  local PSE_WA_1 = p[ 0.000,-0.400, 0.300, 0.000, 0.000, 0.000]
  local PSE_WA_2 = p[-0.300,-0.300, 0.300, 0.000, 0.000, d2r(-90)]
  local PSE_WA_3 = p[-0.300, 0.300, 0.300, 0.000, 0.000, d2r(-135)]
  local PSE_WA_4 = p[ 0.300, 0.300, 0.300, 0.000, 0.000, d2r(135)]
  local PSE_WA_5 = p[ 0.300,-0.300, 0.300, 0.000, 0.000, d2r(90)]
  local PSE_WA_6 = p[ 0.000,-0.600, 0.300, 0.000, 0.000, 0.000]       # reserved
  local PSE_WA_7 = p[ 0.000, 0.000, 0.000, 0.000, 0.000, 0.000]       # reserved
  local PSE_WA_8 = p[ 0.000, 0.000, 0.000, 0.000, 0.000, 0.000]       # reserved
  local PSE_WA_9 = p[ 0.000, 0.000, 0.000, 0.000, 0.000, 0.000]       # reserved
  local PSE_WA_10 = p[ 0.000, 0.000, 0.000, 0.000, 0.000, 0.000]      # reserved

  local JNT_HOME = [-1.22921,-1.29807,-1.79972,-1.6152, 1.57367, 3.48142]
  local JNT_STANDARD_C1 = [ 1.57,-1.57, 1.57,-1.57,-1.57,0]
  local JNT_STANDARD_C2 = [-1.57,-1.57,-1.57,-1.57, 1.57,0]
  local YAW_MIN_DEG = -110
  local YAW_MAX_DEG = 110
  local DISTANCE_TO_CLEARANCE = 0.300
  local RADIUS_HELPER_POSES = 0.300
  local RADIUS_TRANSITION_POSES = 0.400
  local workareas = [WORKAREA_1, WORKAREA_2, WORKAREA_3, WORKAREA_4, WORKAREA_5, WORKAREA_6, WORKAREA_7, WORKAREA_8, WORKAREA_9, WORKAREA_10]
  local poses = [PSE_WA_1, PSE_WA_2, PSE_WA_3, PSE_WA_4, PSE_WA_5, PSE_WA_6, PSE_WA_7, PSE_WA_8, PSE_WA_9, PSE_WA_10]

  ######################### end of adjustment #########################

  local pi = 3.14159265
  local axis_config_current = 0
  local axis_config_new = 0
  local workarea_current = 0
  local workarea_new = 0
  global reverse_rotation = False
  local pose_start = struct(crt = p[0,0,0,0,0,0], jnt = [0,0,0,0,0,0], q = [0,0,0,0,0,0], yaw_too_base = 0.0)
  local pose_help = struct(crt = p[0,0,0,0,0,0], jnt = [0,0,0,0,0,0], q = [0,0,0,0,0,0], yaw_too_base = 0.0)
  local pose_target = struct(crt = p[0,0,0,0,0,0], jnt = [0,0,0,0,0,0], q = [0,0,0,0,0,0], yaw_too_base = 0.0)
  local pose = struct(crt = p[0,0,0,0,0,0], jnt = [0,0,0,0,0,0], q = [0,0,0,0,0,0], yaw_too_base = 0.0)

  def get_tool_free_pose(pose_ref=get_actual_tcp_pose(), dir=[0,0,0], move_in_base_frame=False):
      # get a recovery pose
      # dir is providing the direction and distance in X, Y and Z
      # if 'move_in_base_frame' is set, dir will be interpreted as absolute values for a movement in base frame

      local pose_target = pose_ref
      local i = 0

      if (move_in_base_frame):
          while (i<3):
              # move only,
              # if the demanded position is bigger than zero and the current position is below the demanded one or
              # if the demanded position is smaller than zero and the current position is above the demanded one
              if ((dir[i]>0 and pose_ref[i]<dir[i]) or (dir[i]<0 and pose_ref[i]>dir[i])):
                  pose_target[i] = dir[i]
              end
              i = i + 1
          end
      else:
          pose_target = pose_trans(pose_ref, p[dir[0], dir[1], dir[2], 0, 0, 0])
      end

      return pose_target
  end

  def check_workarea(reference_pose):
      # the actual TCP position is compared to predefined areas (cubic) to determine in which area the robot arm is
      # a workarea is defined as a list of coordinates, where the first 3 values are X, Y, and Z with the smallest values and
      # the next 3 values specify X, Y and Z for the biggest values

      local data_size = size(workareas)
      local i = 0
      local size_workarea = p[0,0,0,0,0,0]
      local pose_workarea = p[0,0,0,0,0,0]

      while (i < data_size[0]):
          pose_workarea = pose_trans(inv(p[workareas[i, 0], workareas[i, 1], workareas[i, 2], 0, 0, 0]), reference_pose)
          size_workarea = pose_sub(p[workareas[i, 3], workareas[i, 4], workareas[i, 5], 0, 0, 0], p[workareas[i, 0], workareas[i, 1], workareas[i, 2], 0, 0, 0])
          if  ((pose_workarea[0]>0 and pose_workarea[0]<size_workarea[0]) and
              (pose_workarea[1]>0 and pose_workarea[1]<size_workarea[1]) and
              (pose_workarea[2]>0 and pose_workarea[2]<size_workarea[2])):
              return i + 1
          end
          i = i + 1
      end
      return 0
  end

  def check_current_axis_config():
      # function determnines, if the arm is oriented in one or the other configuration.
      # it means, that the ellbow joint is flipped and so are the wrist joints.

      local jnt_current = get_actual_joint_positions()

      # ellbow has positiv angle
      if (jnt_current[2]> 0):
          return 1
      # ellbow has negativ angle
      elif (jnt_current[2]< 0):
          return 2
      # angle is 0
      else:
          return 0
      end
  end

  def switch_axis_config(axis_config):
      # function to switch betwwen the axis configuration 1 and 2.

      if (axis_config == 1):
          return 2
      elif (axis_config ==2):
          return 1
      end
  end

  def get_transition_pose_by_workarea(workarea, axis_config):
      # get the correspondig pose from the list of poses

      pose.crt = poses[workarea-1]
      pose.yaw_too_base = get_yaw_too_base(pose.crt)
      pose.q = get_actual_joint_positions()

      if get_inverse_kin_has_solution(pose.crt, qnear=pose.q):
          pose.jnt = get_inverse_kin(pose.crt, qnear=pose.q)
      else:
          popup("no solution found for the transition pose", blocking= True)
      end

      return pose
  end

  def get_transition_pose_by_reference_pose(ref, radius, axis_config):
      # get the correspondig pose from the list of poses

      pose.yaw_too_base = get_yaw_too_base(ref)
      pose.q = get_actual_joint_positions()

      # get coordinates of the circle with the same angle as the given pose to the
      if ref == p[0,0,0,0,0,0]:
          pose.q = JNT_HOME
          pose.jnt = JNT_HOME
          pose.crt = get_forward_kin(pose.jnt)
          return pose
      else:
          pose.crt = p[
              radius * cos(pose.yaw_too_base-pi/2),
              radius * sin(pose.yaw_too_base-pi/2),
              DISTANCE_TO_CLEARANCE,
              0,
              0,
              pose.yaw_too_base + get_locked_yaw()]
      end

      if get_inverse_kin_has_solution(pose.crt, qnear=pose.q):
          pose.jnt = get_inverse_kin(pose.crt, qnear=pose.q)
      else:
          popup("no solution found for the transition pose", blocking= True)
      end

      return pose
  end

  def get_transition_pose_by_yaw(yaw, radius, axis_config):

      pose.yaw_too_base = yaw
      pose.q = get_actual_joint_positions()
      pose.crt = p[
          radius * cos(yaw-pi/2),
          radius * sin(yaw-pi/2),
          DISTANCE_TO_CLEARANCE,
          0,
          0,
          yaw + get_locked_yaw()]

      if get_inverse_kin_has_solution(pose.crt, qnear=pose.q):
          pose.jnt = get_inverse_kin(pose.crt, qnear=pose.q)
      else:
          popup("no solution found for the transition pose", blocking= True)
      end

      return pose
  end

  def get_rounded_mm(value):
      if (value < 0):
          return ceil(value*1000)
      elif (value >= 0):
          return floor(value*1000)
      end
  end

  def get_yaw_too_base(pose):
      # get the yaw relative to the base frame
      local pose_x_mm = 0
      local pose_y_mm = 0
      local yaw = 0

      pose_x_mm = get_rounded_mm(pose[0])
      pose_y_mm = get_rounded_mm(pose[1])

      if (pose_x_mm == 0 and pose_y_mm < 0):
          yaw = 0
      elif (pose_x_mm == 0 and pose_y_mm > 0):
          yaw = pi
      elif (pose_x_mm < 0 and pose_y_mm == 0):
          yaw = -pi/2
      elif (pose_x_mm > 0 and pose_y_mm == 0):
          yaw = pi/2
      else:
          yaw = atan2(pose[0], pose[1])
          if (-pi < yaw) and (yaw < 0):
              yaw = - yaw - pi
          elif (0 < yaw) and (yaw < pi):
              yaw = - yaw + pi
          end
      end
      return yaw
  end

  def adjust_axis_rotation(pose):

      if (0 > pose.yaw_too_base) and (pose.yaw_too_base > d2r(YAW_MIN_DEG)):
          if (pose.jnt[0] > JNT_HOME[0]):
              # calculated axis angle is in the wrong value range
              if axis_config_current == 1:
                  pose.q[0] = JNT_STANDARD_C1[0]
              elif axis_config_current == 2:
                  pose.q[0] = JNT_STANDARD_C2[0]
              end
              reverse_rotation = True
          end
      elif (0 < pose.yaw_too_base) and (pose.yaw_too_base < d2r(YAW_MAX_DEG)):
          if (pose.jnt[0] < JNT_HOME[0]):
              if axis_config_current == 1:
                  pose.q[0] = JNT_STANDARD_C1[0]
              elif axis_config_current == 2:
                  pose.q[0] = JNT_STANDARD_C2[0]
              end
              reverse_rotation = True
          end
      elif (pose.jnt[0] < -2 * pi):
          if axis_config_current == 1:
              pose.q[0] = JNT_STANDARD_C1[0]
          elif axis_config_current == 2:
              pose.q[0] = JNT_STANDARD_C2[0]
          end
          reverse_rotation = True
      elif (pose.jnt[0] > 2 * pi):
          if axis_config_current == 1:
              pose.q[0] = JNT_STANDARD_C1[0]
          elif axis_config_current == 2:
              pose.q[0] = JNT_STANDARD_C2[0]
          end
          reverse_rotation = True
      end
      return pose.q[0]
  end

  def adjust_transition_poses(pose_identifier, keep_rxry=False):
      # adjust the orientation of the transition poses by determining the the current orientation

      local pose_current = get_actual_tcp_pose()
      local jnt_current = get_actual_joint_positions()
      local rpy_current = rotvec2rpy([pose_current[3],pose_current[4],pose_current[5]])
      local rotvec_new = [0,0,0]

      if (pose_identifier == "start"):
          pose = pose_start
      elif (pose_identifier == "target"):
          pose = pose_target
          pose.q[0] = adjust_axis_rotation(pose)
      elif (pose_identifier == "helper"):
          pose = pose_help
      end

      if keep_rxry:
          rotvec_new = rpy2rotvec([rpy_current[0], rpy_current[1], pose.yaw_too_base + get_locked_yaw()])
          pose.crt = p[pose.crt[0], pose.crt[1], pose.crt[2], rotvec_new[0], rotvec_new[1], rotvec_new[2]]

          # adjust preferred joint angles ot the current ones
          pose.q[3] = jnt_current[3]
          pose.q[4] = jnt_current[4]
          pose.q[5] = jnt_current[5]
      end

      if get_inverse_kin_has_solution(pose.crt, qnear=pose.q) and is_within_safety_limits(pose.crt):
          pose.jnt = get_inverse_kin(pose.crt, qnear=pose.q)
      else:
          popup(str_cat("no solution for ", pose_identifier), error=True, blocking=True)
      end
      return pose.jnt
  end

  def get_locked_yaw():
      local pose_current = get_actual_tcp_pose()
      local rpy_current = rotvec2rpy([pose_current[3],pose_current[4],pose_current[5]])
      local rotvec_new = rpy2rotvec([rpy_current[0], rpy_current[1], get_yaw_too_base(pose_current)])
      local pose_reference = p[pose_current[0], pose_current[1], pose_current[2], rotvec_new[0], rotvec_new[1], rotvec_new[2]]
      local pose_to_reference = pose_trans(pose_inv(pose_reference), pose_current)

      return pose_to_reference[5]
  end

  def get_helper_yaw():
      local yaw = 0

      yaw = (pose_start.yaw_too_base + pose_target.yaw_too_base) / 2

      if reverse_rotation and
          ((pose_start.yaw_too_base < 0 and
          pose_target.yaw_too_base < 0) or
          (pose_start.yaw_too_base > 0 and
          pose_target.yaw_too_base > 0)):
            yaw = flip_yaw(yaw)
      elif (pose_start.yaw_too_base < 0 and
            pose_start.yaw_too_base < d2r(YAW_MIN_DEG)) and
            (pose_target.yaw_too_base > 0 and
            pose_target.yaw_too_base > d2r(YAW_MAX_DEG)):
              yaw = flip_yaw(yaw)
      elif (pose_start.yaw_too_base > 0 and
            pose_start.yaw_too_base > d2r(YAW_MAX_DEG)) and
            (pose_target.yaw_too_base < 0 and
            pose_target.yaw_too_base < d2r(YAW_MIN_DEG)):
              yaw = flip_yaw(yaw)
      end
      return yaw
  end

  def flip_yaw(yaw):
      # flips the given yaw 180 degree around
      if (yaw < 0):
          return yaw + pi
      elif (yaw > 0):
          return yaw - pi
      end
  end

  def clear_poses():
      pose = struct(crt = p[0,0,0,0,0,0], jnt = [0,0,0,0,0,0], q = [0,0,0,0,0,0], yaw_too_base = 0.0)
      pose_start = struct(crt = p[0,0,0,0,0,0], jnt = [0,0,0,0,0,0], q = [0,0,0,0,0,0], yaw_too_base = 0.0)
      pose_help = struct(crt = p[0,0,0,0,0,0], jnt = [0,0,0,0,0,0], q = [0,0,0,0,0,0], yaw_too_base = 0.0)
      pose_target = struct(crt = p[0,0,0,0,0,0], jnt = [0,0,0,0,0,0], q = [0,0,0,0,0,0], yaw_too_base = 0.0)
  end

  def do_transition(reference_pose=p[0,0,0,0,0,0], mode=2, keep_rxry=False, a=1.4, v=1.05, r=0.100):
      # the robot will evaluate the current and target workarea
      # after that, the robot will move between the workareas automatically.
      # parameters:
      # reference_pose:   a pose/frame were the robot should work next. If nothing is given, base frame will be used as target
      # keep_rxry:        if true, the robot will keep the orientation of the tool during the movement

      ################# checking #################
      axis_config_current = check_current_axis_config()           # 0: unknown, 1: config 1, 2: config 2
      workarea_current = check_workarea(get_actual_tcp_pose())    # between 0 and the amount of defined workareas
      workarea_new = check_workarea(reference_pose)               # between 0 and the amount of defined workareas
      reverse_rotation = False

      if (workarea_current != 0 and workarea_new != 0) and (workarea_current != workarea_new) or (reference_pose == p[0,0,0,0,0,0]):
          ################# get axisvalues #################
          if (mode == 1):
              pose_start = get_transition_pose_by_workarea(workarea_current, axis_config_current)
              pose_target = get_transition_pose_by_workarea(workarea_new, axis_config_current)
          elif (mode == 2):
              pose_start = get_transition_pose_by_reference_pose(get_actual_tcp_pose(), RADIUS_TRANSITION_POSES, axis_config_current)
              pose_target = get_transition_pose_by_reference_pose(reference_pose, RADIUS_TRANSITION_POSES, axis_config_current)
          end

          global A_Start = pose_start.crt
          global A_End = pose_target.crt
          global A_Start_Yaw = r2d(pose_start.yaw_too_base)
          global A_End_Yaw = r2d(pose_target.yaw_too_base)
          global A_Start_JNT_1 = r2d(pose_start.jnt[0])
          global A_End_JNT_1 = r2d(pose_target.jnt[0])
          global A_Start_JNT = pose_start.jnt
          global A_End_JNT = pose_target.jnt
          global A_Help = pose_help.crt
          global A_Help_Yaw = r2d(pose_help.yaw_too_base)
          global A_Help_JNT = r2d(pose_help.jnt[0])
          # sleep(2)

          ################# adjustments #################
          pose_start.jnt = adjust_transition_poses("start", keep_rxry)
          pose_target.jnt = adjust_transition_poses("target", keep_rxry)

          global A_Start = pose_start.crt
          global A_End = pose_target.crt
          global A_Start_Yaw = r2d(pose_start.yaw_too_base)
          global A_End_Yaw = r2d(pose_target.yaw_too_base)
          global A_Start_JNT_1 = r2d(pose_start.jnt[0])
          global A_End_JNT_1 = r2d(pose_target.jnt[0])
          global A_Start_JNT = pose_start.jnt
          global A_End_JNT = pose_target.jnt

          if (pose_start.crt[1] < 0 and pose_target.crt[1] > 0) or (pose_start.crt[1] > 0 and pose_target.crt[1] < 0):
              pose_help = get_transition_pose_by_yaw(get_helper_yaw(), RADIUS_HELPER_POSES, axis_config_current)
              pose_help.jnt = adjust_transition_poses("helper", keep_rxry)
          end

          global A_Help = pose_help.crt
          global A_Help_Yaw = r2d(pose_help.yaw_too_base)
          global A_Help_JNT = r2d(pose_help.jnt[0])
          global A_Dis_S_H = point_dist(pose_start.crt, pose_help.crt)
          global A_Dis_H_T = point_dist(pose_help.crt, pose_target.crt)
          global A_Dis_S_T = point_dist(pose_start.crt, pose_target.crt)
          # sleep(2)

          ################# movements #################
          if (pose_help.jnt != [0,0,0,0,0,0]):
              if point_dist(get_actual_tcp_pose(), pose_start.crt) > r and point_dist(pose_start.crt, pose_help.crt) > r:
                  movej(pose_start.jnt, a=a, v=v, r=r)
                  if (point_dist(pose_start.crt, pose_help.crt) > r) and (point_dist(pose_target.crt, pose_help.crt) > r):
                      movej(pose_help.jnt, a=a, v=v, r=r)
                  end
              end
          else:
              if point_dist(get_actual_tcp_pose(), pose_start.crt) > r and point_dist(pose_start.crt, pose_target.crt) > r:
                  movej(pose_start.jnt, a=a, v=v, r=r)
              end
          end
          movej(pose_target.jnt, a=a, v=v)
      else:
          # define error
      end

      ################# checking #################
      axis_config_current = check_current_axis_config()           # 0: unknown, 1: config 1, 2: config 2
      workarea_current = check_workarea(get_actual_tcp_pose())    # between 0 and the amount of defined workareas
      clear_poses()
  end
  $ 4 "Script: SCRIPT Utility V5.3.script"
  #*****************************************************
  # customer          :   tbd
  # project name      :   tbd
  #****************************************************
  # controller        :
  # software          :
  #****************************************************
  # author            :   P. Koehnke (+49 1628859904; p.koehnke@unitedrobotics.group)
  # Copyright (c)     :   United Robotics Group Health and Food GmbH
  #                       An der Riede 2
  #                       28816 Stuhr
  #                       Germany
  #****************************************************
  # description       :   utility programs for the application
  # version:      	:   3.1
  # created           :   30.01.2023
  # updated           :
  #****************************************************
  # modifications     :   get_tool_free_pose_2(), get_index_from_list()
  #
  # date              :   05.01.2024
  # name              :   PK
  # reason            :
  #****************************************************

  def found_in_matrix(data, req_id, req_idx):
      local id = -1
      local dimensions = size(data)
      local loop_dataset = 0

      while (id != req_id and loop_dataset < dimensions[0]):
          id = data[loop_dataset, 0]
          if (id == req_id):
              return data[loop_dataset, req_idx]
          else:
              loop_dataset = loop_dataset + 1
          end
      end
  end

  def found_in_list(value, list):
      local idx = 0

      while (idx < length(list)):
          if (value == list[idx]):
              return True
          end
          idx = idx + 1
      end
      return False
  end

  def get_index_from_list(list, value = -1):
      local idx = 0

      while (idx < length(list)):
          if (value == -1):
              if (list[idx] != 0):
                  return idx
              end
          else:
              if (list[idx] == value):
                  return idx
              end
          end
          idx = idx + 1
      end
      return -1
  end

  def pose_RPY2RotVec(pose):
      local rotvec = rpy2rotvec([d2r(pose[3]), d2r(pose[4]), d2r(pose[5])])
      return p[pose[0], pose[1], pose[2], rotvec[0], rotvec[1], rotvec[2]]
  end

  def pose_RotVec2RPY(pose):
      local rpy = rotvec2rpy([pose[3], pose[4], pose[5]])
      return p[pose[0], pose[1], pose[2], r2d(rpy[0]), r2d(rpy[1]), r2d(rpy[2])]
  end

  def swivel(frame_ref, angles = [0, 0, 0], pose = p[0, 0, 0, 0, 0, 0]):

      local rpy_ref = [0, 0, 0]
      local rpy_new = [0, 0, 0]
      local rotvec_new = [0, 0, 0]
      local pose_from = p[0, 0, 0, 0, 0, 0]
      local pose_to = p[0, 0, 0, 0, 0, 0]
      local i = 0

      if (pose == p[0, 0, 0, 0, 0, 0]):
          pose_to = pose_trans(pose_inv(frame_ref), get_actual_tcp_pose())
      else:
          pose_to = pose
      end

      rpy_ref = rotvec2rpy(frame_ref[3], frame_ref[4], frame_ref[5])

      while (i < 3):
          rpy_new[i] = rpy_ref[i] + d2r(angles[i])
          i = i + 1
      end

      rotvec_new = rpy2rotvec(rpy_new)
      pose_from = p[0, 0, 0, rotvec_new[0], rotvec_new[1], rotvec_new[2]]
      pose_to = p[pose_to[0], pose_to[1], pose_to[2], rotvec_new[0], rotvec_new[1], rotvec_new[2]]

      return pose_trans(pose_from, pose_to)
  end

  def get_random_pose(pose_ref, mode = "", range_max = [0, 0, 0]):
      # modi: "cubic", "rotation"
      # getting a random pose in the x/y-plane. range can be set for each
      # translation and rotation.
      local rpy_random = [0, 0, 0]
      local rotvec_random = [0, 0, 0]
      local pose_random = pose_ref
      local i = 0

      if (mode == "cubic"):
          # cubic mode: random pose takes only x, y and z
          i = 0
          while (i < 3):
              pose_random[i] = pose_ref[i] + range_max[i] * (random() - 0.5)
              i = i + 1
          end
          return pose_random

      elif (mode == "rotation"):
          i = 0
          while (i < 3):
              rpy_random[i] = d2r(range_max[i]) * (random() - 0.5)
              i = i + 1
          end
          rotvec_random = rpy2rotvec(rpy_random)
          pose_random = pose_trans(p[0, 0, 0, rotvec_random[0], rotvec_random[1], rotvec_random[2]], pose_ref)
          return pose_random

      else:
          # unknown mode, return pose_ref
          return pose_ref
      end
  end

  def get_pattern_pos_rectangle(counter, direction, pattern, patterninc = [0, 0], patternsize = [0, 0]):
      # defines the position inside a rectangular pattern
      # pattern describes, how many objects are in x-direction and how many in y-direction [x, y]
      # patternsize will give the total length of each direction [x, y]
      local X_Fac = 0
      local Y_Fac = 0
      local max = pattern[0] * pattern[1]
      local i = 0

      if (1 > counter or counter > max):
          counter = 1
      end

      if pattern[0] == 0:
          pattern[0] = 1
      end

      if pattern[1] == 0:
          pattern[1] = 1
      end

      if (direction == "Y" or direction == "y"):
          X_Fac = floor((counter - 1) / pattern[1])
          Y_Fac = (counter - 1) % pattern[1]
      elif (direction == "X" or direction == "x"):
          X_Fac = (counter - 1) % pattern[0]
          Y_Fac = floor((counter - 1) / pattern[0])
      end

      if patternsize != [0, 0]:
          while i < 2:
              if pattern[i] > 1:
                  patterninc[i] = patternsize[i] / (pattern[i] - 1)
              end
              i = i + 1
          end
      end

      return p[X_Fac * patterninc[0], Y_Fac * patterninc[1], 0, 0, 0, 0]
  end

  def get_pattern_pos_circle(counter, radius, angle, direction, pattern, patternsize = [0, 0]):
      # get the patternpos for a circular pattern through a counter
      # need the radius and the angle in radiants
      local X_Fac = 0
      local Y_Fac = 0
      local rad_bow = 0
      local radius_cal = 0
      local ref = p[0, 0, 0, 0, 0, 0]

      if pattern[0] == 0:
          pattern[0] = 1
      end

      if pattern[1] == 0:
          pattern[1] = 1
      end

      if (direction == "Y" or direction == "y"):
          X_Fac = floor((counter - 1) / pattern[1])
          Y_Fac = (counter - 1) % pattern[1]
      elif (direction == "X" or direction == "x"):
          X_Fac = (counter - 1) % pattern[0]
          Y_Fac = floor((counter - 1) / pattern[0])
      end

      # the opening angle will be calculated in x-direction
      # works only between -90 and 90 degree
      if pattern[0] > 1:
          rad_bow = - angle / (pattern[0] - 1) * X_Fac + angle / 2
      end

      if (counter % 2 == 0 and pattern[1] > 1):
          radius_cal = radius - patternsize[1] / (pattern[1])
      else:
          radius_cal = radius + patternsize[1] / (pattern[1])
      end
      ref = p[0, radius_cal, 0, 0, 0, 0]

      return p[ref[0] * cos(rad_bow) - ref[1] * sin(rad_bow), (ref[0] * sin(rad_bow) + ref[1] * cos(rad_bow)) - radius, 0, 0, 0, 0]
  end

  def get_pattern_counter(pose, direction, pattern, patterninc = [0, 0], patternsize = [0, 0]):
      # returns the counter for a pattern from a given cartesian pose
      local patternpose = p[pose[0], pose[1], 0, 0, 0, 0]
      local X_Fac = 0
      local Y_Fac = 0
      local i = 0

      if patternsize != [0, 0]:
          while i < 2:
              if pattern[i] > 1:
                  patterninc[i] = patternsize[i] / (pattern[i] - 1)
              else:
                  pattern[i] = 0
              end
              i = i + 1
          end
      end

      # calculation of the counter in the desired axis-direction
      if (direction == "x" or direction == "X"):
          if patterninc[0] > 0:
              X_Fac = ceil((patternpose[0] + patterninc[0] / 2) / patterninc[0])
              if X_Fac < 0:
                  X_Fac = 0
              end
          end
          if patterninc[1] > 0:
              Y_Fac = floor((patternpose[1] + patterninc[1] / 2) / patterninc[1])
              if Y_Fac < 0:
                  Y_Fac = 0
            end
          end
          return Y_Fac * pattern[0] + X_Fac
      elif (direction == "y" or direction == "Y"):
          if patterninc[0] > 0:
              X_Fac = floor((patternpose[0] + patterninc[0] / 2) / patterninc[0])
          end
          if patterninc[1] > 0:
              Y_Fac = ceil((patternpose[1] + patterninc[1] / 2) / patterninc[1])
          end
          return X_Fac * pattern[1] + Y_Fac
      end
  end

  def get_plc_reg(mod_sig_name):
      return integer_to_binary_list(modbus_get_signal_status(mod_sig_name))
  end

  def set_plc_reg(mod_sig_name, mod_sig_list):
      modbus_set_output_register(mod_sig_name, binary_list_to_integer(mod_sig_list), False)
  end

  def check_decapping(offset = 0, timeout = 5, abort = False):
      # checken, ob der Deckel schon ab ist
      local start = get_actual_tcp_pose()
      local current_offset = 0
      local timecounter = 0
      while (current_offset < offset and not abort):
          current_offset = pose_dist(start, get_actual_tcp_pose())
          timecounter = timecounter + 1
          if (timecounter * 0.5 == timeout):
              break
          end
          sleep(0.5)
      end
      stopl(0.5)
  end

  def check_capping(torque = 0):
      # checken, wann der Deckel verschraubt ist
      force_mode(get_actual_tcp_pose(), [0, 0, 1, 0, 0, 0], [0, 0, -2.0, 0, 0, 0], 2, [0, 0, 0.100, 0, 0, 0])
  end

  def is_reachable(frame, poses, offsets = [0, 0, 0]):
      local idx = 0
      local pose = p[0, 0, 0, 0, 0, 0]

      while (idx < length(poses)):
          pose = poses[idx]
          pose[0] = pose[0] + offsets[0]
          pose[1] = pose[1] + offsets[1]
          pose[2] = pose[2] + offsets[2]

          if pose != p[0, 0, 0, 0, 0, 0]:
              if (not get_inverse_kin_has_solution(pose_trans(frame, pose))):
                  textmsg(str_cat(str_cat("Pose ", to_str(idx + 1)), " is not reachable"))
                  return False
              end
          end
          idx = idx + 1
      end
      return True
  end

  def is_within_limits(frame, poses, offsets = [0, 0, 0]):
      local idx = 0
      local pose = p[0, 0, 0, 0, 0, 0]

      while (idx < length(poses)):
          pose = poses[idx]
          pose[0] = pose[0] + offsets[0]
          pose[1] = pose[1] + offsets[1]
          pose[2] = pose[2] + offsets[2]

          if is_reachable(frame = frame, poses = poses, offsets = offsets):
              if (not is_within_safety_limits(get_inverse_kin(pose_trans(frame, pose), get_actual_joint_positions()))):
                  textmsg(str_cat(str_cat("Pose ", to_str(idx + 1)), "is out of joint limits"))
                  return False
              else:
                  idx = idx + 1
              end
          else:
              return False
          end
      end
      return True
  end
  $ 5 "Script: SCRIPT Vision Config V0.2.script"
  CAM_LM = struct(id=0, type="", size=0, related_itm=0, capture_relation="")
  global CAM_Result = make_list(0, 0, 50)

  def create_landmark(id=0, type="", size=0, related_itm=0, capture_relation=""):
      return struct(id=id, type=type, size=size, related_itm=related_itm, capture_relation=capture_relation)
  end


  CAM_LMs = [
    create_landmark(id=1, type="aruco_7x7", size=0.1, related_itm=1, capture_relation="front_right"),
    create_landmark(id=4, type="aruco_7x7", size=0.1, related_itm=2, capture_relation="straight_left"),
    create_landmark(id=3, type="aruco_7x7", size=0.1, related_itm=2, capture_relation="straight_left"),
    create_landmark(id=8, type="aruco_7x7", size=0.1, related_itm=2, capture_relation="right"),
    create_landmark(id=5, type="aruco_7x7", size=0.1, related_itm=5, capture_relation="left"),
    create_landmark(id=6, type="aruco_7x7", size=0.1, related_itm=2, capture_relation="straight_left")
  ]

  CAM_Capture_Poses = struct(
    front_left = p[0.350,-0.330,0.500,0.353,-0.323,-1.458],
    left = p[0.350,0.000,0.500,0.353,-0.323,-1.458],
    back_left = p[0.350,0.220,0.500,0.353,-0.323,-1.458],
    back_right = p[-0.350,0.000,0.500,0.579,0.240,0.760],
    right = p[-0.350,-0.300,0.500,0.206,0.206,1.561],
    front_right = p[-0.350,-0.400,0.500,0.242,0.903,2.480],
    straight_left = p[0.375,-0.000,0.500,0.815,-0.815,-1.412],
    front = p[0,0,0,0,0,0]
  )

  def get_capture_pose(lm):
      if (lm.capture_relation == "front_left"):
          return CAM_Capture_Poses.front_left
      elif (lm.capture_relation == "left"):
          return CAM_Capture_Poses.left
      elif (lm.capture_relation == "back_left"):
          return CAM_Capture_Poses.back_left
      elif (lm.capture_relation == "back_right"):
          return CAM_Capture_Poses.back_right
      elif (lm.capture_relation == "right"):
          return CAM_Capture_Poses.right
      elif (lm.capture_relation == "straight_left"):
         return CAM_Capture_Poses.straight_left
      else:
          # error
          return get_actual_tcp_pose()
      end
  end
  $ 6 "Script: 001 SCRIPT Errors and Warnings Deifnes V0.2.script"

  #*****************************************************
  # customer          :   UK Essen
  # project name      :   P1132
  #****************************************************
  # controller        :
  # software          :
  #****************************************************
  # author            :   E.Petrichenko
  # Copyright (c)     :   United Robotics Group Health and Food GmbH
  #                       An der Riede 2
  #                       28816 Stuhr
  #                       Germany
  #****************************************************
  # description       :   centrifuge actions for the application
  # version:      	:   0.1
  # created           :   22.08.2024
  # updated           :
  #****************************************************
  # modifications     :
  #
  # date              :
  # name              :
  # reason            :
  #****************************************************


  #################################### VARIABLES DEFINITIONS ###################################

  ERROR_POSE_NOT_REACHABLE = 1002
  ERROR_ROBOT_ARM_NOT_IN_HOME_POSE = 1006
  ERROR_NO_OBJECT_TO_PICK = 1010
  ERROR_NOT_DOCKED = 2003
  ERROR_NOT_REACHABLE_TARGET = 2007
  ERROR_CHARGING_NOT_STARTED = 2008
  ERROR_AMR_WRONG_MODE = 2009
  ERROR_UNKNOWN_POSE = 2010
  ERROR_NO_LANDMARK = 3002
  ERROR_WRONG_ORDER = 4002
  ERROR_CENTRIFUGE_CONNECTION = 5001
  ERROR_CENTRIFUGE_POWER = 5002
  ERROR_CENTRIFUGE = 5003
  ERROR_CENTRIFUGE_LID = 5004
  ERROR_CANNOT_OPEN_HATCH = 5006
  ERROR_CANNOT_CLOSE_HATCH = 5008
  ERROR_CANNOT_ROTATE = 5010
  ERROR_CANNOT_START = 5011
  ERROR_WRONG_KEY_POSE = 5012
  ERROR_MISSIING_CENTRACK = 5013

  WARNING_POSE_NOT_REACHABLE = 1002
  WARNING_BATTERY_LEVEL = 2002
  WARNING_NOT_REACHABLE_TARGET = 2007


  ERROR = struct(
      FLAG = False,
      ID = 0,
      MSG = "")

  WARNING = struct(
      FLAG = False,
      ID = 0,
      MSG = "")


  #################################### FUNCTIONS ###################################

  def set_error(error_id):
      ERROR.ID = error_id
      if (ERROR.ID == 0):
          ERROR.FLAG = False
          ERROR.MSG = ""
      else:
          ERROR.FLAG = True
          if(ERROR.ID == ERROR_POSE_NOT_REACHABLE):
              ERROR.MSG = "Pose is not reachable"
          elif(ERROR.ID == ERROR_NO_OBJECT_TO_PICK):
              ERROR.MSG = "No object to pick"
          elif(ERROR.ID == ERROR_NO_LANDMARK):
              ERROR.MSG = "No landmark detected"
          elif(ERROR.ID == ERROR_ROBOT_ARM_NOT_IN_HOME_POSE):
              ERROR.MSG = "Robot arm cannot go to home pose"
          elif(ERROR.ID == ERROR_AMR_WRONG_MODE):
              ERROR.MSG = "AMR is in the wrong mode"
          elif(ERROR.ID == ERROR_NOT_DOCKED):
              ERROR.MSG = "Could not dock to the charger"
          elif(ERROR.ID == ERROR_NOT_REACHABLE_TARGET):
              ERROR.MSG = "Could not reach the target"
          elif(ERROR.ID == ERROR_CHARGING_NOT_STARTED):
              ERROR.MSG = "Could not start charging"
          elif(ERROR.ID == ERROR_UNKNOWN_POSE):
              ERROR.MSG = "Unknown navigation target"
          elif(ERROR.ID == ERROR_CANNOT_OPEN_HATCH):
              ERROR.MSG = "Centrifuge Cannot open the hatch"
          elif(ERROR.ID == ERROR_CENTRIFUGE_CONNECTION):
              ERROR.MSG = "Cannot reach centrifuge"
          elif (ERROR.ID == ERROR_CANNOT_CLOSE_HATCH):
              ERROR.MSG = "Centrifuge Cannot close the hatch"
          elif (ERROR.ID == ERROR_CANNOT_START):
              ERROR.MSG = "Centrifuge Cannot start"
          elif (ERROR.ID == ERROR_CANNOT_ROTATE):
              ERROR.MSG = "Centrifuge Cannot rotate the rotor"
          elif (ERROR.ID == ERROR_WRONG_ORDER):
              ERROR.MSG = "Wrong parameter was recieved"
          elif (ERROR.ID == ERROR_CENTRIFUGE):
              ERROR.MSG = "Centrifuge is in Error"
          elif (ERROR.ID == ERROR_WRONG_KEY_POSE):
              ERROR.MSG = "Key is in the wrong position"
          elif(ERROR.ID == ERROR_MISSIING_CENTRACK):
              ERROR.MSG = "Missing rack for centrifuge set"
          elif(ERROR.ID == ERROR_CENTRIFUGE_POWER):
              ERROR.MSG = "Centrifuge is turned off"
          elif(ERROR.ID == ERROR_CENTRIFUGE_LID):
              ERROR.MSG = "Lid of the centrifuge is opened"
          else:
              ERROR.MSG = "Unknown code"
          end
          textmsg("ERROR:",ERROR)
      end
  end

  def set_warning(warning_id):
      WARNING.ID = warning_id
      if (WARNING.ID == 0):
          WARNING.FLAG = False
          WARNING.MSG = ""
      else:
          WARNING.FLAG = True
          if(WARNING.ID == WARNING_POSE_NOT_REACHABLE):
              WARNING.MSG = "Pose is not reachable"
          elif(WARNING.ID == WARNING_BATTERY_LEVEL):
              WARNING.MSG = "Batery level dropped to a certain level"
          elif(WARNING.ID == WARNING_NOT_REACHABLE_TARGET):
              WARNING.MSG = "Not reachable location of AMR"
          else:
              WARNING.MSG = "Unknown code"
          end
          textmsg("WARNING:",WARNING)
      end
  end


  def reset_error():
    ERROR.ID = 0
    ERROR.FLAG = False
    ERROR.MSG = ""
  end


  def reset_warning():
      WARNING.ID = 0
      WARNING.FLAG = False
      WARNING.MSG = ""
    end
  $ 46 "reset_error()"
  reset_error()
  $ 47 "Action≔131"
  global Action=131
  $ 48 "ITM_ID≔1"
  global ITM_ID=1
  $ 49 "JIG≔7"
  global JIG=7
  $ 50 "CMD_Stop≔ False "
  global CMD_Stop=  False
  $ 51 "PSE_T≔get_actual_tcp_pose()"
  global PSE_T= get_actual_tcp_pose ()
  $ 52 "MoveJ"
  $ 53 "PSE_T" "breakAfter"
  movej(PSE_T, a=1.3962634015954636, v=1.0471975511965976)
  $ 54 "Set"
  set_tcp(p[0.0,0.0,0.161,3.1415,0.0,0.0])
  $ 55 "Robot Program"
  $ 56 "PreSettings"
  $ 57 "CAM_LM_Detected≔ False "
  global CAM_LM_Detected=  False
  $ 58 "CAM_Captures≔0"
  global CAM_Captures=0
  $ 59 "CAM_Pose≔p[0,0,0,0,0,0]"
  global CAM_Pose=p[0,0,0,0,0,0]
  $ 60 "CAM_LM_Refinmnt≔ False "
  global CAM_LM_Refinmnt=  False
  $ 61 "CAM_LM_Refined≔ False "
  global CAM_LM_Refined=  False
  $ 62 "CAM_LM_Deviatn≔p[0,0,0,0,0,0]"
  global CAM_LM_Deviatn=p[0,0,0,0,0,0]
  $ 63 "CAM_LM_ID≔0"
  global CAM_LM_ID=0
  $ 64 "CAM_Done≔ False "
  global CAM_Done=  False
  $ 65 "CAM_CNT_Obj≔0"
  global CAM_CNT_Obj=0
  $ 66 "CAM_Result = []"
  CAM_Result = []
  $ 67 "OBJ_Detected≔ False "
  global OBJ_Detected=  False
  $ 68 "FRM_Reference≔p[0,0,0,0,0,0]"
  global FRM_Reference=p[0,0,0,0,0,0]
  $ 69 "'=========='"
  # '=========='
  $ 70 "Switch Action"
  switch_1 = Action
  $ 71 "Case 13"
  if (13 == switch_1):
  elif (15 == switch_1):
    $ 189 "Case 15"
  elif (131 == switch_1):
    $ 235 "Case 131"
    $ 236 "Read (SensoPart)"
    $ 237 "Action_Info≔'search for landmark'"
    global Action_Info="search for landmark"
    $ 238 "CAM_LM≔CAM_LMs[ITM_ID-1]"
    global CAM_LM=CAM_LMs[ITM_ID-1]
    $ 239 "CAM_Relation≔CAM_LM.capture_relation"
    global CAM_Relation=CAM_LM.capture_relation
    $ 240 "go to capture pose"
    $ 243 "If ITM_ID≟1 and JIG≟7"
    if (ITM_ID == 1  and  JIG == 7):
      $ 244 "PSE_T≔ULM_Cap_SSRack"
      global PSE_T=ULM_Cap_SSRack
    else:
      $ 245 "ElseIf ITM_ID≟5 and JIG≟7"
      if (ITM_ID == 5  and  JIG == 7):
        $ 246 "PSE_T≔FRM_Cap_SSTable"
        global PSE_T=FRM_Cap_SSTable
      end
    end
    $ 247 "do_transition(PSE_T, keep_rxry=False)"
    do_transition(PSE_T, keep_rxry=False)
    $ 248 "Set"
    set_tcp(p[0.0,0.0,0.161,3.1415,0.0,0.0])
    $ 249 "MoveJ"
    $ 250 "PSE_T" "breakAfter"
    movej(PSE_T, a=1.3962634015954636, v=1.7453292519943295)
    $ 251 "CAM_Pose≔get_actual_tcp_pose()"
    global CAM_Pose= get_actual_tcp_pose ()
    $ 252 "Loop  not CAM_Done and  not ERROR.FLAG and  not CMD_Stop"
    while (  not  CAM_Done  and    not  ERROR.FLAG  and    not  CMD_Stop):
      $ 253 "adjust capture pose"
      $ 254 "If CAM_LM_Detected and CAM_LM_Refinmnt"
      if (CAM_LM_Detected  and  CAM_LM_Refinmnt):
        $ 255 "PSE_T≔p[0,0,0.300,0,0,0]"
        global PSE_T=p[0,0,0.300,0,0,0]
        $ 256 "CAM_Pose≔PSE_T"
        global CAM_Pose=PSE_T
        $ 257 "If  not is_reachable(FRM_Reference,[PSE_T])"
        if (  not  is_reachable(FRM_Reference,[PSE_T])):
          $ 258 "Error"
          $ 259 "set_error(ERROR_POSE_NOT_REACHABLE)"
          set_error(ERROR_POSE_NOT_REACHABLE)
        end
        $ 260 "If  not ERROR.FLAG"
        if (  not  ERROR.FLAG):
          $ 261 "MoveJ"
          $ 262 "PSE_T" "breakAfter"
          set_tcp(p[0.0,0.0,0.161,0.0,0.0,0.0])
          movej(pose_trans(FRM_Reference, PSE_T), a=0.8726646259971648, v=1.3962634015954636)
          $ 263 "CAM_LM_Refined≔ True "
          global CAM_LM_Refined=  True
        end
      else:
        $ 264 "ElseIf  not CAM_LM_Detected and CAM_Captures>0"
        if (  not  CAM_LM_Detected  and  CAM_Captures>0):
          $ 265 "MoveL"
          $ 266 "If FRM_Reference≟p[0,0,0,0,0,0]"
          if (FRM_Reference == p[0,0,0,0,0,0]):
            $ 267 "PSE_T≔get_random_pose(pose_ref=CAM_Pose, mode='cubic', range_max=[0.150,0.150,0.020])"
            global PSE_T=get_random_pose(pose_ref=CAM_Pose, mode="cubic", range_max=[0.150,0.150,0.020])
          else:
            $ 268 "Else" "noBreak"
            $ 269 "PSE_T≔get_random_pose(pose_ref=CAM_Pose, mode='rotation', range_max=[10,10,0])"
            global PSE_T=get_random_pose(pose_ref=CAM_Pose, mode="rotation", range_max=[10,10,0])
            $ 270 "CAM_LM_Refined≔ True "
            global CAM_LM_Refined=  True
          end
          $ 271 "If get_inverse_kin_has_solution(pose_trans(FRM_Reference, PSE_T))"
          if (get_inverse_kin_has_solution( pose_trans (FRM_Reference, PSE_T))):
            $ 272 "PSE_T" "breakAfter"
            set_tcp(p[0.0,0.0,0.161,0.0,0.0,0.0])
            movel(pose_trans(FRM_Reference, PSE_T), a=0.03, v=0.05)
          else:
            $ 273 "Else" "noBreak"
            $ 274 "'If random pose is out of reach, set the initial cam pose'"
            # 'If random pose is out of reach, set the initial cam pose'
            $ 275 "PSE_T≔CAM_Pose"
            global PSE_T=CAM_Pose
          end
        end
      end
      $ 276 "Wait: 2.0"
      sleep(2.0)
      $ 277 "trigger"
      # begin: URCap Program Node
      #   Source: SensoPart VISOR Robotic, 2.0.0, SensoPart Industriesensorik GmbH
      #   Type: VISOR Trigger
      $ 278 "# 1 VISOR Trigger"
      visor_changeJob(1, "Landmark Detection", 3000)
      visor_trigger(1, 3000, "arm")
      # end: URCap Program Node
      $ 279 "CAM_LM_Deviatn≔visor_getPose3d(1, 0)"
      global CAM_LM_Deviatn= visor_getPose3d (1, 0)
      $ 280 "If CAM_LM_Deviatn≠PSE_Z"
      if (CAM_LM_Deviatn != PSE_Z):
        $ 281 "CAM_LM_Detected≔ True "
        global CAM_LM_Detected=  True
        $ 282 "CAM_Captures≔0"
        global CAM_Captures=0
      else:
        $ 283 "Else" "noBreak"
        $ 284 "CAM_LM_Detected≔ False "
        global CAM_LM_Detected=  False
        $ 285 "CAM_Captures≔CAM_Captures+1"
        global CAM_Captures=CAM_Captures+1
      end
      $ 286 "result"
      $ 287 "If CAM_LM_Detected"
      if (CAM_LM_Detected):
        $ 288 "If (CAM_LM_Refinmnt and CAM_LM_Refined) or  not CAM_LM_Refinmnt"
        if ((CAM_LM_Refinmnt  and  CAM_LM_Refined)  or    not  CAM_LM_Refinmnt):
          $ 346 "If ITM_ID≟1 and JIG≟7"
          if (ITM_ID == 1  and  JIG == 7):
            $ 354 "ULM_SS_Rack≔pose_trans(CAM_LM_Deviatn, ULM_SS_Rack)"
            global ULM_SS_Rack= pose_trans (CAM_LM_Deviatn, ULM_SS_Rack)
          else:
            $ 356 "ElseIf ITM_ID≟5 and JIG≟7"
            if (ITM_ID == 5  and  JIG == 7):
              $ 358 "FRM_SS_SSTable[0]=CAM_LM_Deviatn[0]"
              FRM_SS_SSTable[0]=CAM_LM_Deviatn[0]
              $ 359 "FRM_SS_SSTable[1]=CAM_LM_Deviatn[1]"
              FRM_SS_SSTable[1]=CAM_LM_Deviatn[1]
            end
          end
          $ 360 "CAM_Done≔ True "
          global CAM_Done=  True
        end
      else:
        $ 361 "ElseIf  not CAM_LM_Detected and CAM_Captures<CAM_PRM_Retries"
        if (  not  CAM_LM_Detected  and  CAM_Captures<CAM_PRM_Retries):
          $ 362 "CAM_LM_Refined≔ False "
          global CAM_LM_Refined=  False
        else:
          $ 363 "ElseIf CAM_Captures≥CAM_PRM_Retries"
          if (CAM_Captures >= CAM_PRM_Retries):
            $ 364 "CAM_Done≔ True "
            global CAM_Done=  True
            $ 365 "Error"
            $ 366 "set_error(ERROR_NO_LANDMARK)"
            set_error(ERROR_NO_LANDMARK)
          end
        end
      end
    end
  elif (151 == switch_1):
    $ 367 "Case 151"
    $ 368 "Detect (SensoPart)"
    $ 369 "go to capture pose"
    $ 370 "FRM_Reference≔ULM_Input"
    global FRM_Reference=ULM_Input
    $ 372 "PSE_T≔ULM_Cap_SSRack"
    global PSE_T=ULM_Cap_SSRack
    $ 373 "do_transition(pose_trans(FRM_Reference, PSE_T), keep_rxry=False)"
    do_transition( pose_trans (FRM_Reference, PSE_T), keep_rxry=False)
    $ 374 "JNT_Q≔get_actual_joint_positions()"
    global JNT_Q= get_actual_joint_positions ()
    $ 375 "JNT_Q≔[JNT_Q[0], JNT_Q[1], JNT_Q[2], JNT_Q[3], JNT_Q[4], 0]"
    global JNT_Q=[JNT_Q[0], JNT_Q[1], JNT_Q[2], JNT_Q[3], JNT_Q[4], 0]
    $ 376 "Set"
    set_tcp(p[0.0,0.0,0.161,0.0,0.0,0.0])
    $ 377 "movej(get_inverse_kin(pose_trans(FRM_Reference, PSE_T), qnear=JNT_Q))"
    movej(get_inverse_kin( pose_trans (FRM_Reference, PSE_T), qnear=JNT_Q))
    $ 378 "CAM_Pose≔pose_trans(pose_inv(FRM_Reference), get_actual_tcp_pose())"
    global CAM_Pose= pose_trans ( pose_inv (FRM_Reference),  get_actual_tcp_pose ())
    $ 379 "Loop  not CAM_Done and  not ERROR.FLAG and  not CMD_Stop"
    while (  not  CAM_Done  and    not  ERROR.FLAG  and    not  CMD_Stop):
      $ 380 "If  not OBJ_Detected and CAM_Captures>0"
      if (  not  OBJ_Detected  and  CAM_Captures>0):
        $ 381 "MoveL"
        $ 382 "If FRM_Reference≟p[0,0,0,0,0,0]"
        if (FRM_Reference == p[0,0,0,0,0,0]):
          $ 384 "PSE_T≔get_random_pose(pose_ref=CAM_Pose, mode='rotation', range_max=[15,15,0])"
          global PSE_T=get_random_pose(pose_ref=CAM_Pose, mode="rotation", range_max=[15,15,0])
        else:
          $ 385 "Else" "noBreak"
          $ 386 "PSE_T≔get_random_pose(pose_ref=CAM_Pose, mode='rotation', range_max=[10,10,0])"
          global PSE_T=get_random_pose(pose_ref=CAM_Pose, mode="rotation", range_max=[10,10,0])
        end
        $ 387 "If get_inverse_kin_has_solution(pose_trans(FRM_Reference, PSE_T))"
        if (get_inverse_kin_has_solution( pose_trans (FRM_Reference, PSE_T))):
          $ 388 "PSE_T" "breakAfter"
          set_tcp(p[0.0,0.0,0.161,0.0,0.0,0.0])
          movel(pose_trans(FRM_Reference, PSE_T), a=0.03, v=0.05)
        else:
          $ 389 "Else" "noBreak"
          $ 390 "'If random pose is out of reach, set the initial cam pose'"
          # 'If random pose is out of reach, set the initial cam pose'
          $ 391 "PSE_T≔CAM_Pose"
          global PSE_T=CAM_Pose
          $ 392 "PSE_T" "breakAfter"
          set_tcp(p[0.0,0.0,0.161,0.0,0.0,0.0])
          movel(pose_trans(FRM_Reference, PSE_T), a=0.03, v=0.05)
        end
      end
      $ 393 "Wait: 0.5"
      sleep(0.5)
      $ 394 "Set"
      set_tcp(p[0.0,0.0,0.161,3.1415,0.0,0.0])
      # begin: URCap Program Node
      #   Source: SensoPart VISOR Robotic, 2.0.0, SensoPart Industriesensorik GmbH
      #   Type: VISOR Trigger
      $ 395 "# 1 VISOR Trigger"
      visor_changeJob(1, "Object Detection Single", 3000)
      visor_trigger(1, 3000, "arm")
      # end: URCap Program Node
      $ 396 "If visor_isResponseOk(1)"
      if ( visor_isResponseOk (1)):
        $ 397 "CAM_CNT_Obj≔visor_partsFound(1)"
        global CAM_CNT_Obj= visor_partsFound (1)
        $ 398 "CAM_OBJ_Pose≔visor_getPose3d(1, 0)"
        global CAM_OBJ_Pose= visor_getPose3d (1, 0)
        $ 399 "If CAM_CNT_Obj>0"
        if (CAM_CNT_Obj>0):
          $ 400 "CAM_OBJ_Color≔visor_getAdditionalData(1, 0)"
          global CAM_OBJ_Color= visor_getAdditionalData (1, 0)
          $ 401 "CAM_DetectScore≔to_num(visor_getAdditionalData(1, 1))/1000"
          global CAM_DetectScore=to_num( visor_getAdditionalData (1, 1))/1000
          $ 402 "OBJ_Detected≔ True "
          global OBJ_Detected=  True
        end
      else:
        $ 403 "Else" "noBreak"
        $ 404 "CAM_Captures≔CAM_Captures+1"
        global CAM_Captures=CAM_Captures+1
      end
      $ 405 "If OBJ_Detected"
      if (OBJ_Detected):
        $ 406 "Get object data"
        $ 407 "PRC_CntDetect≔0"
        global PRC_CntDetect=0
        $ 408 "Loop PRC_CntDetect<CAM_CNT_Obj"
        while (PRC_CntDetect<CAM_CNT_Obj):
          $ 409 "get object and jig number"
          $ 410 "If ITM_ID≟1 and JIG≟7"
          if (ITM_ID == 1  and  JIG == 7):
            $ 411 "FRM_Reference≔ULM_Cap_SSRack"
            global FRM_Reference=ULM_Cap_SSRack
          else:
            $ 412 "ElseIf ITM_ID≟5 and JIG≟7"
            if (ITM_ID == 5  and  JIG == 7):
              $ 413 "FRM_Reference≔FRM_Cap_SSTable"
              global FRM_Reference=FRM_Cap_SSTable
            end
          end
          $ 416 "PSE_T≔pose_trans(pose_inv(FRM_Reference), CAM_OBJ_Pose)"
          global PSE_T= pose_trans ( pose_inv (FRM_Reference), CAM_OBJ_Pose)
          $ 417 "CAM_Result.append(get_pattern_counter(PSE_T, 'X', pattern=[10, 5], patternsize=[0.181, 0.081]))"
          CAM_Result.append(get_pattern_counter(PSE_T, "X", pattern=[10, 5], patternsize=[0.181, 0.081]))
          $ 419 "PRC_CntDetect≔PRC_CntDetect+1"
          global PRC_CntDetect=PRC_CntDetect+1
        end
        $ 420 "CAM_Done≔ True "
        global CAM_Done=  True
      else:
        $ 421 "ElseIf CAM_Captures≥CAM_PRM_Retries"
        if (CAM_Captures >= CAM_PRM_Retries):
          $ 422 "CAM_Done≔ True "
          global CAM_Done=  True
        else:
          $ 423 "Else" "noBreak"
          $ 424 "CAM_Captures≔CAM_Captures+1"
          global CAM_Captures=CAM_Captures+1
        end
      end
    end
  end
  $ 425 "'=========='"
  # '=========='
  $ 426 "PostSettings"
  $ 427 "FRM_Reference≔p[0,0,0,0,0,0]"
  global FRM_Reference=p[0,0,0,0,0,0]
  $ 428 "Set"
  set_tcp(p[0.0,0.0,0.161,3.1415,0.0,0.0])
  $ 429 "CAM_Pose≔p[0,0,0,0,0,0]"
  global CAM_Pose=p[0,0,0,0,0,0]
  $ 430 "Action≔0"
  global Action=0
  $ 431 "Action_Info≔''"
  global Action_Info=""
end
